(* IEC 61131-3 sources: Palletizer_Control_with_Automation_Studio/Palletizer/Logical/Libraries/MTBasics, 3 files *)

(* ---- MTBasics.typ ---- *)
TYPE
	MTBasicsDT1InternalType : 	STRUCT  (*Internal variables of function block MTBasicsDT1.*)
		CycleTime : REAL; (*Task cycle time. Unit: [µs].*)
		ParametersValid : BOOL; (*Data for internal use.*)
		Gain : REAL; (*Data for internal use.*)
		TimeConstant : REAL; (*Data for internal use.*)
		Numerator : ARRAY[0..1]OF LREAL; (*Data for internal use.*)
		Denominator : ARRAY[0..1]OF LREAL; (*Data for internal use.*)
		BVector : ARRAY[0..1]OF LREAL; (*Data for internal use.*)
		AVector : ARRAY[0..1]OF LREAL; (*Data for internal use.*)
		XVector : ARRAY[0..1]OF LREAL; (*Data for internal use.*)
		PresetOK : BOOL; (*Data for internal use.*)
		PresetCoefficients : LREAL; (*Data for internal use.*)
		InOld : REAL; (*Data for internal use.*)
		UpdateOld : BOOL; (*Data for internal use.*)
		EnableOld : BOOL; (*Data for internal use.*)
		EnableDone : BOOL; (*Data for internal use.*)
		DisabledBusy : BOOL; (*Data for internal use.*)
		CounterOld : UDINT; (*Data for internal use.*)
		SysRefParaNew : BOOL; (*Data for internal use.*)
		SystemReference : MTTransferFcnType; (*Data for internal use.*)
	END_STRUCT;
	MTBasicsDT2InternalType : 	STRUCT  (*Internal variables of function block MTBasicsDT2.*)
		CycleTime : REAL; (*Task cycle time. Unit: [µs].*)
		ParametersValid : BOOL; (*Data for internal use.*)
		Gain : REAL; (*Data for internal use.*)
		TimeConstant1 : REAL; (*Data for internal use.*)
		TimeConstant2 : REAL; (*Data for internal use.*)
		Numerator : ARRAY[0..2]OF LREAL; (*Data for internal use.*)
		Denominator : ARRAY[0..2]OF LREAL; (*Data for internal use.*)
		BVector : ARRAY[0..2]OF LREAL; (*Data for internal use.*)
		AVector : ARRAY[0..2]OF LREAL; (*Data for internal use.*)
		XVector : ARRAY[0..1]OF LREAL; (*Data for internal use.*)
		PresetOK : BOOL; (*Data for internal use.*)
		PresetCoefficients : LREAL; (*Data for internal use.*)
		InOld : REAL; (*Data for internal use.*)
		UpdateOld : BOOL; (*Data for internal use.*)
		EnableOld : BOOL; (*Data for internal use.*)
		EnableDone : BOOL; (*Data for internal use.*)
		DisabledBusy : BOOL; (*Data for internal use.*)
		CounterOld : UDINT; (*Data for internal use.*)
		SysRefParaNew : BOOL; (*Data for internal use.*)
		SystemReference : MTTransferFcnType; (*Data for internal use.*)
	END_STRUCT;
	MTBasicsIntegratorInternalType : 	STRUCT  (*Internal variables of function block MTBasicsIntegrator.*)
		CycleTime : REAL; (*Task cycle time. Unit: [s].*)
		ParametersValid : BOOL; (*Data for internal use.*)
		Gain : REAL; (*Data for internal use.*)
		BVector : ARRAY[0..1]OF LREAL; (*Data for internal use.*)
		AVector : ARRAY[0..1]OF LREAL; (*Data for internal use.*)
		XVector : LREAL; (*Data for internal use.*)
		OutPresetValue : REAL; (*Data for internal use.*)
		SetOutOld : BOOL; (*Data for internal use.*)
		UpdateOld : BOOL; (*Data for internal use.*)
		EnableOld : BOOL; (*Data for internal use.*)
		EnableDone : BOOL; (*Data for internal use.*)
		DisabledBusy : BOOL; (*Data for internal use.*)
		CounterOld : UDINT; (*Data for internal use.*)
		SysRefParaNew : BOOL; (*Data for internal use.*)
		SystemReference : MTTransferFcnType; (*Data for internal use.*)
	END_STRUCT;
	MTBasicsLevelCtrlInternalType : 	STRUCT  (*Internal variables of function block MTBasicsLevelController.*)
		CycleTime : REAL; (*Task cycle time. Unit: [s].*)
		ParametersValid : BOOL; (*Data for internal use.*)
		Parameter : MTBasicsLevelCtrlParType; (*Data for internal use.*)
		State : USINT; (*Data for internal use.*)
		UpdateOld : BOOL; (*Data for internal use.*)
		EnableOld : BOOL; (*Data for internal use.*)
	END_STRUCT;
	MTBasicsLevelCtrlParType : 	STRUCT  (*Level controller parameters.*)
		OutputValue1 : REAL; (*1st Output value.*)
		OutputValue2 : REAL; (*2nd Output value.*)
		OutputValue3 : REAL; (*3rd Output value.*)
		ThresholdLevel1 : REAL; (*Threshold level from OutputValue2 to OutputValue1.*)
		ThresholdLevel2 : REAL; (*Threshold level from OutputValue1 to OutputValue2.*)
		ThresholdLevel3 : REAL; (*Threshold level from OutputValue3 to OutputValue2.*)
		ThresholdLevel4 : REAL; (*Threshold level from OutputValue2 to OutputValue3.*)
	END_STRUCT;
	MTBasicsLimiterInternalType : 	STRUCT  (*Internal variables of function block MTBasicsLimiter.*)
		CycleTime : REAL; (*Task cycle time. Unit: [s].*)
		ParametersValid : BOOL; (*Data for internal use.*)
		MaxOut : REAL; (*Data for internal use.*)
		MinOut : REAL; (*Data for internal use.*)
		MaxPosSlewRate : REAL; (*Data for internal use.*)
		MaxNegSlewRate : REAL; (*Data for internal use.*)
		Out : REAL; (*Data for internal use.*)
		OutOld : REAL; (*Data for internal use.*)
		UpperOutLimit : REAL; (*Data for internal use.*)
		LowerOutLimit : REAL; (*Data for internal use.*)
		SetOutOld : BOOL; (*Data for internal use.*)
		UpdateOld : BOOL; (*Data for internal use.*)
		EnableOld : BOOL; (*Data for internal use.*)
	END_STRUCT;
	MTBasicsOscTuningInternalType : 	STRUCT  (*Internal variables of function block MTBasicsOscillationTuning.*)
		CycleTime : REAL; (*Task cycle time. Unit: [s].*)
		ParametersValid : BOOL; (*Data for internal use.*)
		State : USINT; (*State of tuning.*)
		CriticalGain : REAL; (*Critical gain.*)
		OscillationPeriod : REAL; (*Period of oscillation.*)
		NumberOfOscillations : USINT; (*Number of osscilations.*)
		NumberOfPhases : USINT; (*Number of current tuning phase.*)
		MaxRelayOut : REAL; (*Lower limit for output during tuning.*)
		MinRelayOut : REAL; (*Upper limit for output during tuning.*)
		SetValue : REAL; (*Data for internal use.*)
		AverageOutValue : REAL; (*Data for internal use.*)
		MaxActValueTime : ARRAY[0..3]OF REAL; (*Data for internal use.*)
		MinActValueTime : ARRAY[0..3]OF REAL; (*Data for internal use.*)
		MaxActValue : ARRAY[0..3]OF REAL; (*Data for internal use.*)
		MinActValue : ARRAY[0..3]OF REAL; (*Data for internal use.*)
		TuningTime : REAL; (*Data for internal use.*)
		StartingActValue : REAL; (*Data for internal use.*)
		ControlError : REAL; (*Data for internal use.*)
		ActValueAverageAmplitude : REAL; (*Data for internal use.*)
		AverageActValue : REAL; (*Data for internal use.*)
		AverageMaxActValue : REAL; (*Data for internal use.*)
		AverageMinActValue : REAL; (*Data for internal use.*)
		AmplitudeRatio : REAL; (*Data for internal use.*)
		DeltaOut : REAL; (*Data for internal use.*)
		EffectiveDirection : SINT; (*Data for internal use.*)
		StartOld : BOOL; (*Data for internal use.*)
		MinOscillationAmplitude : REAL; (*Data for internal use.*)
		MinOut : REAL; (*Data for internal use.*)
		MaxOut : REAL; (*Data for internal use.*)
		TemporaryQuality : REAL; (*Data for internal use.*)
		TemporaryDerivativeTime : REAL; (*Data for internal use.*)
		TemporaryIntegrationTime : REAL; (*Data for internal use.*)
		TemporaryGain : REAL; (*Data for internal use.*)
		Update : BOOL; (*Data for internal use.*)
		UpdateOld : BOOL; (*Data for internal use.*)
		EnableOld : BOOL; (*Data for internal use.*)
		AverageOutValueSum : REAL; (*Data for internal use.*)
		AverageTime : LREAL; (*Data for internal use.*)
	END_STRUCT;
	MTBasicsPFMInternalType : 	STRUCT  (*Internal variables of function block MTBasicsPFM.*)
		CycleTime : REAL; (*Task cycle time. Unit: [s].*)
		ParametersValid : BOOL; (*Data for internal use.*)
		In : REAL; (*Data for internal use.*)
		PulseWidth : REAL; (*Data for internal use.*)
		MinPause : REAL; (*Data for internal use.*)
		Area : REAL; (*Data for internal use.*)
		AreaC : REAL; (*Data for internal use.*)
		OffTime : REAL; (*Data for internal use.*)
		OnTime : REAL; (*Data for internal use.*)
		Update : BOOL; (*Data for internal use.*)
		UpdateOld : BOOL; (*Data for internal use.*)
		EnableOld : BOOL; (*Data for internal use.*)
	END_STRUCT;
	MTBasicsPIDInternalType : 	STRUCT  (*Internal variables of function block MTBasicsPID.*)
		CycleTime : REAL; (*Task cycle time. Unit: [s].*)
		ParametersValid : BOOL; (*Data for internal use.*)
		PIDParameters : MTPIDParametersType; (*Data for internal use.*)
		MinOut : REAL; (*Data for internal use.*)
		MaxOut : REAL; (*Data for internal use.*)
		Invert : BOOL; (*Data for internal use.*)
		ControlError : REAL; (*Data for internal use.*)
		ControlErrorOld : REAL; (*Data for internal use.*)
		Out : REAL; (*Data for internal use.*)
		HoldIntegration : MTPIDIntegrationEnum; (*Data for internal use.*)
		IntegrationPartPresetValue : REAL; (*Data for internal use.*)
		SetIntegrationPart : BOOL; (*Data for internal use.*)
		SetIntegrationPartOld : BOOL; (*Data for internal use.*)
		EnableTrackingOld : BOOL; (*Data for internal use.*)
		PID_StatusID : DINT; (*Data for internal use.*)
		UpdateOld : BOOL; (*Data for internal use.*)
		EnableOld : BOOL; (*Data for internal use.*)
		EnableDone : BOOL; (*Data for internal use.*)
		DisabledBusy : BOOL; (*Data for internal use.*)
		CounterOld : UDINT; (*Data for internal use.*)
		SysRefParaNew : BOOL; (*Data for internal use.*)
		SystemReference : MTTransferFcnType; (*Data for internal use.*)
	END_STRUCT;
	MTBasicsPT1InternalType : 	STRUCT  (*Internal variables of function block MTBasicsPT1.*)
		CycleTime : REAL; (*Task cycle time. Unit: [s].*)
		ParametersValid : BOOL; (*Data for internal use.*)
		Gain : REAL; (*Data for internal use.*)
		TimeConstant : REAL; (*Data for internal use.*)
		Numerator : ARRAY[0..1]OF LREAL; (*Data for internal use.*)
		Denominator : ARRAY[0..1]OF LREAL; (*Data for internal use.*)
		BVector : ARRAY[0..1]OF LREAL; (*Data for internal use.*)
		AVector : ARRAY[0..1]OF LREAL; (*Data for internal use.*)
		XVector : ARRAY[0..1]OF LREAL; (*Data for internal use.*)
		OutPresetValue : REAL; (*Data for internal use.*)
		PresetCoefficients : LREAL; (*Data for internal use.*)
		PresetOK : BOOL; (*Data for internal use.*)
		SetOutOld : BOOL; (*Data for internal use.*)
		UpdateOld : BOOL; (*Data for internal use.*)
		EnableOld : BOOL; (*Data for internal use.*)
		EnableDone : BOOL; (*Data for internal use.*)
		DisabledBusy : BOOL; (*Data for internal use.*)
		CounterOld : UDINT; (*Data for internal use.*)
		SysRefParaNew : BOOL; (*Data for internal use.*)
		SystemReference : MTTransferFcnType; (*Data for internal use.*)
	END_STRUCT;
	MTBasicsPT2InternalType : 	STRUCT  (*Internal variables of function block MTBasicsPT2.*)
		CycleTime : REAL; (*Task cycle time. Unit: [µs].*)
		ParametersValid : BOOL; (*Data for internal use.*)
		Gain : REAL; (*Data for internal use.*)
		TimeConstant1 : REAL; (*Data for internal use.*)
		TimeConstant2 : REAL; (*Data for internal use.*)
		Numerator : ARRAY[0..2]OF LREAL; (*Data for internal use.*)
		Denominator : ARRAY[0..2]OF LREAL; (*Data for internal use.*)
		BVector : ARRAY[0..2]OF LREAL; (*Data for internal use.*)
		AVector : ARRAY[0..2]OF LREAL; (*Data for internal use.*)
		XVector : ARRAY[0..1]OF LREAL; (*Data for internal use.*)
		OutPresetValue : REAL; (*Data for internal use.*)
		PresetCoefficients : LREAL; (*Data for internal use.*)
		PresetOK : BOOL; (*Data for internal use.*)
		SetOutOld : BOOL; (*Data for internal use.*)
		UpdateOld : BOOL; (*Data for internal use.*)
		EnableOld : BOOL; (*Data for internal use.*)
		EnableDone : BOOL; (*Data for internal use.*)
		DisabledBusy : BOOL; (*Data for internal use.*)
		CounterOld : UDINT; (*Data for internal use.*)
		SysRefParaNew : BOOL; (*Data for internal use.*)
		SystemReference : MTTransferFcnType; (*Data for internal use.*)
	END_STRUCT;
	MTBasicsPWMInternalType : 	STRUCT  (*Internal variables of function block MTBasicsPWM.*)
		CycleTime : REAL; (*Task cycle time. Unit: [s].*)
		ParametersValid : BOOL; (*Data for internal use.*)
		Mode : MTBasicsPWMModeEnum; (*Data for internal use.*)
		MinPulseWidth : REAL; (*Data for internal use.*)
		Period : REAL; (*Data for internal use.*)
		In : REAL; (*Data for internal use.*)
		OnTime : REAL; (*Data for internal use.*)
		OffTime : REAL; (*Data for internal use.*)
		PeriodCounter : REAL; (*Data for internal use.*)
		OnTimeCounter : REAL; (*Data for internal use.*)
		UpdateOld : BOOL; (*Data for internal use.*)
		EnableOld : BOOL; (*Data for internal use.*)
	END_STRUCT;
	MTBasicsPWMModeEnum :
		( (*Pulse mode.*)
		mtBASICS_PULSE_BEGINNING := 0, (*Pulse at the beginning of a period.*)
		mtBASICS_PULSE_MIDDLE := 1 (*Pulse in the middle of a period.*)
		);
	MTBasicsPWMScheduleBufferPtrType : 	STRUCT  (*Buffer pointers of the PWMSchedule.*)
		In : REAL; (*Data for internal use.*)
		OnTime1 : REAL; (*Data for internal use.*)
		OnTime2 : REAL; (*Data for internal use.*)
		OffTime1 : REAL; (*Data for internal use.*)
		OffTime2 : REAL; (*Data for internal use.*)
		OnTimeCounter : REAL; (*Data for internal use.*)
	END_STRUCT;
	MTBasicsPWMScheduleBufferType : 	STRUCT  (*Buffer parameters of the PWMSchedule.*)
		ActIndex : UINT; (*Data for internal use.*)
		ActBufferElements : UINT; (*Data for internal use.*)
		OldBufferElements : {REDUND_UNREPLICABLE} UINT; (*Data for internal use.*)
		PointerTimes : REFERENCE TO MTBasicsPWMScheduleBufferPtrType; (*Data for internal use.*)
		PointerOut : REFERENCE TO BOOL; (*Data for internal use.*)
	END_STRUCT;
	MTBasicsPWMScheduleInternalType : 	STRUCT  (*Internal variables of function block MTBasicsPWM.*)
		CycleTime : REAL; (*Task cycle time. Unit: [s].*)
		ParametersValid : BOOL; (*Data for internal use.*)
		NumberOfInputs : UINT; (*Data for internal use.*)
		Mode : MTBasicsPWMScheduleModeEnum; (*Data for internal use.*)
		MinPulseWidth : REAL; (*Data for internal use.*)
		MinPause : REAL; (*Data for internal use.*)
		Period : REAL; (*Data for internal use.*)
		FreeDutyCycle : REAL; (*Data for internal use.*)
		PeriodCounter : REAL; (*Data for internal use.*)
		Buffer : MTBasicsPWMScheduleBufferType; (*Data for internal use.*)
		UpdateOld : BOOL; (*Data for internal use.*)
		EnableOld : {REDUND_UNREPLICABLE} BOOL; (*Data for internal use.*)
		InhibitUpdate : BOOL; (*Data for internal use.*)
		Update : BOOL; (*Data for internal use.*)
		StatusIDUpdate : DINT; (*Data for internal use.*)
	END_STRUCT;
	MTBasicsPWMScheduleModeEnum :
		( (*Schedule mode.*)
		mtBASICS_SHIFT_PULSE := 0, (*Shift the puls.*)
		mtBASICS_SPLIT_PULSE := 1 (*Split the puls.*)
		);
	MTBasicsStepTuningBufElemType : 	STRUCT  (*Buffer element of MTBasicsStepTuning.*)
		TimeIndex : UDINT; (*Data for internal use.*)
		In : LREAL; (*Data for internal use.*)
		IntIn : LREAL; (*Data for internal use.*)
		IntTimeIn : LREAL; (*Data for internal use.*)
		IntTime2In : LREAL; (*Data for internal use.*)
		Int2In : LREAL; (*Data for internal use.*)
		Int3In : LREAL; (*Data for internal use.*)
		TSum : LREAL; (*Data for internal use.*)
		dTSum : LREAL; (*Data for internal use.*)
		d2TSum : LREAL; (*Data for internal use.*)
		dyACD : LREAL; (*Data for internal use.*)
		d2yACD : LREAL; (*Data for internal use.*)
		d3yACD : LREAL; (*Data for internal use.*)
		DiffIn : LREAL; (*Data for internal use.*)
		Diff2In : LREAL; (*Data for internal use.*)
	END_STRUCT;
	MTBasicsStepTuningInternalType : 	STRUCT  (*Internal variables of function block MTBasicsStepTuning.*)
		CycleTime : REAL; (*Task cycle time. Unit: [s].*)
		ParametersValid : BOOL; (*Data for internal use.*)
		MinActValue : REAL; (*Data for internal use.*)
		MaxActValue : REAL; (*Data for internal use.*)
		MaxTuningTime : REAL; (*Data for internal use.*)
		StepHeight : REAL; (*Data for internal use.*)
		State : MTBasicsStepTuningStateEnum; (*Data for internal use.*)
		TuningTime : REAL; (*Data for internal use.*)
		Area : REAL; (*Data for internal use.*)
		StartActValue : REAL; (*Data for internal use.*)
		SumTime : REAL; (*Data for internal use.*)
		PlantGain : REAL; (*Data for internal use.*)
		LQError : REAL; (*Data for internal use.*)
		LQOutput : ARRAY[0..1]OF REAL; (*Data for internal use.*)
		LQParameterVector : ARRAY[0..2]OF REAL; (*Data for internal use.*)
		ActValueOld : REAL; (*Data for internal use.*)
		SystemSettlingTime : REAL; (*Data for internal use.*)
		SettlingIndex : UINT; (*Data for internal use.*)
		NumberOfSettlingValues : UINT; (*Data for internal use.*)
		NoiseDeadBand : REAL; (*Data for internal use.*)
		StartOld : BOOL; (*Data for internal use.*)
		UpdateOld : BOOL; (*Data for internal use.*)
		EnableOld : BOOL; (*Data for internal use.*)
		Slope : REAL; (*Data for internal use.*)
	END_STRUCT;
	MTBasicsStepTuningStateEnum :
		( (*Tuning state.*)
		mtBASICS_STATE_READY := 1, (*The function block waits for a rising edge of Start.*)
		mtBASICS_STATE_SETTLING := 2, (*It is checked, if the system is in an idle state.*)
		mtBASICS_STATE_STEP := 3, (*The output Out is set to the value StepHeight.*)
		mtBASICS_STATE_CALCULATE_PID := 4 (*PID parameters are calculated.*)
		);
	MTBasicsTimeDelayFcnParaType : 	STRUCT  (*Internal variables for time delay function parameters.*)
		DelayCounter : UDINT; (*Data for internal use.*)
		ActBufferIndex : UDINT; (*Data for internal use.*)
		ActBufferElements : UDINT; (*Data for internal use.*)
		OldBufferElements : UDINT; (*Data for internal use.*)
		DelayTimeAct : REAL; (*Data for internal use.*)
		BufferPointer : REFERENCE TO REAL; (*Data for internal use.*)
	END_STRUCT;
	MTBasicsTimeDelayInternalType : 	STRUCT  (*Internal variables of function block MTBasicsTimeDelay.*)
		CycleTime : REAL; (*Task cycle time. Unit: [s].*)
		DelayTime : REAL; (*Data for internal use.*)
		ParametersValid : BOOL; (*Data for internal use.*)
		InitialValue : REAL; (*Data for internal use.*)
		EnableOld : BOOL; (*Data for internal use.*)
		TimeDelayFcnPara : {REDUND_UNREPLICABLE} MTBasicsTimeDelayFcnParaType; (*Data for internal use.*)
	END_STRUCT;
END_TYPE

(* ---- MTBasics.fun ---- *)
{REDUND_OK} FUNCTION_BLOCK MTBasicsDT1 (*First-order derivative action element.*)
	VAR_INPUT
		Enable : BOOL; (*Enables/Disables the function block.*)
		Gain : REAL; (*Gain factor.*)
		TimeConstant : REAL; (*Time constant. Unit: [s]. Valid value range: TimeConstant >= 0.*)
		Update : BOOL; (*Updates the parameters listed above on a rising edge.*)
		In : REAL; (*Input value.*)
	END_VAR
	VAR_OUTPUT
		Busy : BOOL; (*Function block is busy.*)
		Active : BOOL; (*Function block is active.*)
		Error : BOOL; (*Indicates an error.*)
		StatusID : DINT; (*Status information.*)
		UpdateDone : BOOL; (*Update is done.*)
		Out : REAL; (*Output value.*)
		SystemReference : {REDUND_UNREPLICABLE} UDINT; (*System reference.*)
	END_VAR
	VAR
		Internal : MTBasicsDT1InternalType; (*Data for internal use.*)
	END_VAR
END_FUNCTION_BLOCK

{REDUND_OK} FUNCTION_BLOCK MTBasicsDT2 (*Second-order derivative action element.*)
	VAR_INPUT
		Enable : BOOL; (*Enables/Disables the function block.*)
		Gain : REAL; (*Gain factor.*)
		TimeConstant1 : REAL; (*Time constant. Unit: [s]. Valid value range: TimeConstant1 >= 0.*)
		TimeConstant2 : REAL; (*Time constant. Unit: [s]. Valid value range: TimeConstant2 >= 0.*)
		Update : BOOL; (*Updates the parameters listed above on a rising edge.*)
		In : REAL; (*Input value.*)
	END_VAR
	VAR_OUTPUT
		Busy : BOOL; (*Function block is busy.*)
		Active : BOOL; (*Function block is active.*)
		Error : BOOL; (*Indicates an error.*)
		StatusID : DINT; (*Status information.*)
		UpdateDone : BOOL; (*Update is done.*)
		Out : REAL; (*Output value.*)
		SystemReference : {REDUND_UNREPLICABLE} UDINT; (*System reference.*)
	END_VAR
	VAR
		Internal : MTBasicsDT2InternalType; (*Data for internal use.*)
	END_VAR
END_FUNCTION_BLOCK

{REDUND_OK} FUNCTION_BLOCK MTBasicsIntegrator (*Integrator.*)
	VAR_INPUT
		Enable : BOOL; (*Enables/Disables the function block.*)
		Gain : REAL; (*Gain factor. Valid value range: Gain >= 0.*)
		Update : BOOL; (*Updates the parameters listed above on a rising edge.*)
		In : REAL; (*Input value.*)
		OutPresetValue : REAL; (*Preset value for Out output.*)
		SetOut : BOOL; (*Sets Out to OutPresetValue on rising edge.*)
		HoldOut : BOOL; (*Freezes the function block.*)
	END_VAR
	VAR_OUTPUT
		Busy : BOOL; (*Function block is busy.*)
		Active : BOOL; (*Function block is active.*)
		Error : BOOL; (*Indicates an error.*)
		StatusID : DINT; (*Status information.*)
		UpdateDone : BOOL; (*Update is done.*)
		Out : REAL; (*Output value.*)
		SystemReference : {REDUND_UNREPLICABLE} UDINT; (*System reference.*)
	END_VAR
	VAR
		Internal : MTBasicsIntegratorInternalType; (*Data for internal use.*)
	END_VAR
END_FUNCTION_BLOCK

{REDUND_OK} FUNCTION_BLOCK MTBasicsLevelController (*Level controller.*)
	VAR_INPUT
		Enable : BOOL; (*Enables/Disables the function block.*)
		Parameter : MTBasicsLevelCtrlParType; (*3-step controller parameters.*)
		Update : BOOL; (*Updates the parameters listed above on a rising edge.*)
		In : REAL; (*Input value.*)
	END_VAR
	VAR_OUTPUT
		Active : BOOL; (*Function block is active.*)
		Error : BOOL; (*Indicates an error.*)
		StatusID : DINT; (*Status information.*)
		UpdateDone : BOOL; (*Update is done.*)
		Out : REAL; (*Output value.*)
	END_VAR
	VAR
		Internal : MTBasicsLevelCtrlInternalType; (*Data for internal use.*)
	END_VAR
END_FUNCTION_BLOCK

{REDUND_OK} FUNCTION_BLOCK MTBasicsLimiter (*Limiter.*)
	VAR_INPUT
		Enable : BOOL; (*Enables/Disables the function block.*)
		MinOut : REAL; (*Lower output variable limit. Valid value range: MinOut < MaxOut.*)
		MaxOut : REAL; (*Upper output variable limit. Valid value range: MaxOut > MinOut.*)
		MaxPosSlewRate : REAL; (*Maximum output variable ramp for ramp-up. Unit: [1/s]. Valid value range: MaxPosSlewRate >= 0.*)
		MaxNegSlewRate : REAL; (*Maximum output variable ramp for the ramp-down. Unit: [1/s]. Valid value range: MaxNegSlewRate >= 0.*)
		Update : BOOL; (*Updates the parameters listed above on a rising edge.*)
		In : REAL; (*Input value.*)
		OutPresetValue : REAL; (*Preset value for Out output.*)
		SetOut : BOOL; (*Sets Out to OutPresetValue on rising edge.*)
	END_VAR
	VAR_OUTPUT
		Active : BOOL; (*Function block is active.*)
		Error : BOOL; (*Indicates an error.*)
		StatusID : DINT; (*Status information.*)
		UpdateDone : BOOL; (*Update is done.*)
		Out : REAL; (*Output value.*)
	END_VAR
	VAR
		Internal : MTBasicsLimiterInternalType; (*Data for internal use.*)
	END_VAR
END_FUNCTION_BLOCK

{REDUND_OK} FUNCTION_BLOCK MTBasicsOscillationTuning (*Oscillation tuning for PID.*)
	VAR_INPUT
		Enable : BOOL; (*Enables/Disables the function block.*)
		SetValue : REAL; (*Reference variable (setpoint).*)
		MinOut : REAL; (*Lower manipulated variable limit. Valid value range: MinOut < MaxOut.*)
		MaxOut : REAL; (*Upper manipulated variable limit. Valid value range: MaxOut > MinOut.*)
		Invert : BOOL; (*Inverts the direction of the controller.*)
		Update : BOOL; (*Updates the parameters listed above on a rising edge.*)
		ActValue : REAL; (*Actual measured value.*)
		Start : BOOL; (*Starts the tuning (on positive edge).*)
	END_VAR
	VAR_OUTPUT
		Active : BOOL; (*Function block is active.*)
		Error : BOOL; (*Indicates an error.*)
		StatusID : DINT; (*Status information.*)
		UpdateDone : BOOL; (*Update is done.*)
		Out : REAL; (*Output value (manipulated variable). Value range: MinOut <= Out <= MaxOut.*)
		TuningActive : BOOL; (*Tuning is active.*)
		TuningDone : BOOL; (*Tuning completed.*)
		Quality : REAL; (*Quality of the oscillation tuning. Unit: [%]. Value range: 0 (low) ... 100 (high).*)
		PIDParameters : MTPIDParametersType; (*PID parameters.*)
	END_VAR
	VAR
		Internal : MTBasicsOscTuningInternalType; (*Data for internal use.*)
	END_VAR
END_FUNCTION_BLOCK

{REDUND_OK} FUNCTION_BLOCK MTBasicsPFM (*Pulse frequency modulator.*)
	VAR_INPUT
		Enable : BOOL; (*Enables/Disables the function block.*)
		PulseWidth : REAL; (*Pulse width at the output. Unit: [s]. Valid value range: PulseWidth >= task cycle time.*)
		MinPause : REAL; (*Minimum pause between the pulses at the output. Unit: [s]. Valid value range: MinPause >= task cycle time.*)
		Update : BOOL; (*Updates the parameters listed above on a rising edge.*)
		DutyCycle : REAL; (*Input value.*)
	END_VAR
	VAR_OUTPUT
		Active : BOOL; (*Function block is active.*)
		Error : BOOL; (*Indicates an error.*)
		StatusID : DINT; (*Status information.*)
		UpdateDone : BOOL; (*Update is done.*)
		Out : BOOL; (*Output value.*)
	END_VAR
	VAR
		Internal : MTBasicsPFMInternalType; (*Data for internal use.*)
	END_VAR
END_FUNCTION_BLOCK

{REDUND_OK} FUNCTION_BLOCK MTBasicsPID (*PID controller.*)
	VAR_INPUT
		Enable : BOOL; (*Enables/Disables the function block.*)
		PIDParameters : MTPIDParametersType; (*PID parameters.*)
		MinOut : REAL;
		MaxOut : REAL;
		Invert : BOOL;
		Update : BOOL; (*Updates the parameters listed above on a rising edge.*)
		SetValue : REAL; (*Set value (reference variable).*)
		ActValue : REAL; (*Actual value (controlled variable).*)
		IntegrationPartPresetValue : REAL; (*Preset value for the integral component IntegrationPart.*)
		SetIntegrationPart : BOOL; (*A positive edge on SetIntegrationPart sets the integral component IntegrationPart of the PID controller to IntegrationPartPresetValue.*)
		HoldOut : BOOL; (*Freezes the function block.*)
		TrackingValue : REAL; (*Preset value for the integral component IntegrationPart.*)
		EnableTracking : BOOL; (*A positive edge on SetIntegrationPart sets the integral component IntegrationPart of the PID controller to IntegrationPartPresetValue.*)
		HoldIntegration : MTPIDIntegrationEnum; (*PID parameters.*)
	END_VAR
	VAR_OUTPUT
		Busy : BOOL; (*Function block is busy.*)
		Active : BOOL; (*Function block is active.*)
		Error : BOOL; (*Indicates an error.*)
		StatusID : DINT; (*Status information.*)
		UpdateDone : BOOL; (*Update is done.*)
		Out : REAL; (*Controller output. Value range: MinOut <= Out <= MaxOut.*)
		ControlError : REAL; (*Control error.*)
		ProportionalPart : REAL; (*Proportional component.*)
		IntegrationPart : REAL; (*Integral component.*)
		DerivativePart : REAL; (*Derivative component.*)
		TrackingActive : BOOL; (*Derivative component.*)
		IntegrationStatus : MTPIDIntegrationEnum; (*Derivative component.*)
		SystemReference : {REDUND_UNREPLICABLE} UDINT; (*System reference.*)
	END_VAR
	VAR
		Internal : MTBasicsPIDInternalType; (*Data for internal use.*)
	END_VAR
END_FUNCTION_BLOCK

{REDUND_OK} FUNCTION_BLOCK MTBasicsPT1 (*First-order delay element.*)
	VAR_INPUT
		Enable : BOOL; (*Enables/Disables the function block.*)
		Gain : REAL; (*Gain factor.*)
		TimeConstant : REAL; (*Time constant. Unit: [s]. Valid value range: TimeConstant >= 0.*)
		Update : BOOL; (*Updates the parameters listed above on a rising edge.*)
		In : REAL; (*Input value.*)
		OutPresetValue : REAL; (*Preset value for Out output.*)
		SetOut : BOOL; (*Sets Out to OutPresetValue on rising edge.*)
	END_VAR
	VAR_OUTPUT
		Busy : BOOL; (*Function block is busy.*)
		Active : BOOL; (*Function block is active.*)
		Error : BOOL; (*Indicates an error.*)
		StatusID : DINT; (*Status information.*)
		UpdateDone : BOOL; (*Update is done.*)
		Out : REAL; (*Output value.*)
		SystemReference : {REDUND_UNREPLICABLE} UDINT; (*System reference.*)
	END_VAR
	VAR
		Internal : MTBasicsPT1InternalType; (*Data for internal use.*)
	END_VAR
END_FUNCTION_BLOCK

{REDUND_OK} FUNCTION_BLOCK MTBasicsPT2 (*Second-order delay element.*)
	VAR_INPUT
		Enable : BOOL; (*Enables/Disables the function block.*)
		Gain : REAL; (*Gain.*)
		TimeConstant1 : REAL; (*Time constant. Unit: [s]. Valid value range: TimeConstant1 >= 0.*)
		TimeConstant2 : REAL; (*Time constant. Unit: [s]. Valid value range: TimeConstant2 >= 0.*)
		Update : BOOL; (*Updates the parameters listed above on a rising edge.*)
		In : REAL; (*Input value.*)
		OutPresetValue : REAL; (*Preset value for Out output.*)
		SetOut : BOOL; (*Sets Out to OutPresetValue on rising edge.*)
	END_VAR
	VAR_OUTPUT
		Busy : BOOL; (*Function block is busy.*)
		Active : BOOL; (*Function block is active.*)
		Error : BOOL; (*Indicates an error.*)
		StatusID : DINT; (*Status information.*)
		UpdateDone : BOOL; (*Update is done.*)
		Out : REAL; (*Output value.*)
		SystemReference : {REDUND_UNREPLICABLE} UDINT; (*System reference.*)
	END_VAR
	VAR
		Internal : MTBasicsPT2InternalType; (*Data for internal use.*)
	END_VAR
END_FUNCTION_BLOCK

{REDUND_OK} FUNCTION_BLOCK MTBasicsPWM (*Pulse width modulator.*)
	VAR_INPUT
		Enable : BOOL; (*Enables/Disables the function block.*)
		Mode : MTBasicsPWMModeEnum; (*Pulse mode.*)
		MinPulseWidth : REAL; (*Minimum duration of the output actuator pulses and pauses. Unit: [s]. Valid value range: MinPulseWidth < Period.*)
		Period : REAL; (*Period for the output actuator pulses. Unit: [s]. Valid value range: Period > task cycle time.*)
		Update : BOOL; (*Updates the parameters listed above on a rising edge.*)
		DutyCycle : REAL; (*Input value. Unit: [%]. Valid value range: 0 <= DutyCycle <= 100.*)
	END_VAR
	VAR_OUTPUT
		Active : BOOL; (*Function block is active.*)
		Error : BOOL; (*Indicates an error.*)
		StatusID : DINT; (*Status information.*)
		UpdateDone : BOOL; (*Update is done.*)
		Out : BOOL; (*Output value.*)
	END_VAR
	VAR
		Internal : MTBasicsPWMInternalType; (*Data for internal use.*)
	END_VAR
END_FUNCTION_BLOCK

{REDUND_CONTEXT} FUNCTION_BLOCK MTBasicsPWMSchedule (*Multiple pulse width modulator.*)
	VAR_INPUT
		Enable : BOOL; (*Enables/Disables the function block.*)
		Period : REAL; (*Period for the output actuator pulses. Unit: [s]. Permitted range: Period > Task cycle time.*)
		MinPulseWidth : REAL; (*Minimum duration of the pulses. Unit: [s]. Permitted range: Task cycle time <= MinPulseWidth < Period.*)
		MinPause : REAL; (*Minimum duration of the pauses. Unit: [s]. Permitted range: Task cycle time <= MinPause < Period.*)
		Mode : MTBasicsPWMScheduleModeEnum; (*Pulse mode.*)
		Update : BOOL; (*Updates the parameters listed above on a rising edge.*)
		NumberOfInputs : UINT; (*Number of input signals. Permitted range: 0 < NumberOfInputs <= 500.*)
		DutyCycle : {REDUND_UNREPLICABLE} UDINT; (*Address of an array of real with the iput values. Unit of values of the assigned array: [%].*)
	END_VAR
	VAR_OUTPUT
		Active : BOOL; (*Function block is active.*)
		Error : BOOL; (*Indicates an error.*)
		StatusID : DINT; (*Status information.*)
		UpdateDone : BOOL; (*Update is done.*)
		Out : {REDUND_UNREPLICABLE} UDINT; (*Address for an array of bool with the output values.*)
	END_VAR
	VAR
		Internal : MTBasicsPWMScheduleInternalType; (*Data for internal use.*)
	END_VAR
END_FUNCTION_BLOCK

{REDUND_OK} FUNCTION_BLOCK MTBasicsStepTuning (*Step tuning for PID.*)
	VAR_INPUT
		Enable : BOOL; (*Enables/Disables the function block.*)
		SystemSettlingTime : REAL; (*System settling time.*)
		MaxTuningTime : REAL; (*Maximum tuning time*)
		MinActValue : REAL; (*Minimum value of the controlled variable.*)
		MaxActValue : REAL; (*Maximum value of the controlled variable.*)
		Update : BOOL; (*Updates the parameters listed above on a rising edge.*)
		ActValue : REAL; (*Actual measured value.*)
		StepHeight : REAL; (*Height of step to be applied.*)
		Start : BOOL; (*Starts the tuning (on positive edge).*)
	END_VAR
	VAR_OUTPUT
		Active : BOOL; (*Function block is active.*)
		Error : BOOL; (*Indicates an error.*)
		StatusID : DINT; (*Status information.*)
		UpdateDone : BOOL; (*Update is done.*)
		Out : REAL; (*Output value (manipulated variable). Value range: MinOut <= Out <= MaxOut.*)
		TuningActive : BOOL; (*Tuning is active.*)
		TuningDone : BOOL; (*Tuning completed.*)
		PIDParameters : MTPIDParametersType; (*PID parameters.*)
		Quality : REAL; (*Quality of the step tuning. Unit: [%]. Value range: 0 (low) ... 100 (high).*)
		TuningState : MTBasicsStepTuningStateEnum; (*Current state of the tuning procedure.*)
	END_VAR
	VAR
		Internal : MTBasicsStepTuningInternalType; (*Data for internal use.*)
	END_VAR
END_FUNCTION_BLOCK

{REDUND_CONTEXT} FUNCTION_BLOCK MTBasicsTimeDelay (*Delay element.*)
	VAR_INPUT
		Enable : BOOL; (*Enables/Disables the function block.*)
		DelayTime : REAL; (*Delay time. Unit: [s]. Valid value range: 0 <= DelayTime <= "10000 · task cycle time".*)
		In : REAL; (*Input value.*)
		InitialValue : REAL; (*Initial value for Out output.*)
	END_VAR
	VAR_OUTPUT
		Active : BOOL; (*Function block is active.*)
		Error : BOOL; (*Indicates an error.*)
		StatusID : DINT; (*Status information.*)
		Out : REAL; (*Output value.*)
	END_VAR
	VAR
		Internal : MTBasicsTimeDelayInternalType; (*Data for internal use.*)
	END_VAR
END_FUNCTION_BLOCK

(* ---- MTBasics.var ---- *)
(*Error*)
VAR CONSTANT
	mtBCD_ERR_TIME_CONSTANT1_INVALID : DINT := -1058012139; (*Chosen first time constant is invalid.*)
	mtBCD_ERR_TIME_CONSTANT2_INVALID : DINT := -1058012138; (*Chosen second time constant is invalid.*)
	mtBCD_ERR_THRESHOLD_NOT_DEFINED : DINT := -1058012137; (*Chosen values for the threshold levels are invalid.*)
	mtBCD_ERR_THRESHOLD_INVALID : DINT := -1058012136; (*One of the values for the threshold levels is invalid.*)
	mtBCD_ERR_OUT_VALUE_NOT_DEFINED : DINT := -1058012135; (*Chosen output values are invalid.*)
	mtBCD_ERR_OUTPUT_LIMIT_INVALID : DINT := -1058012134; (*Chosen limitations for output are invalid.*)
	mtBCD_ERR_MAX_POS_SLEW_RATE_NEG : DINT := -1058012133; (*Chosen slew rate for positive direction is invalid.*)
	mtBCD_ERR_MAX_NEG_SLEW_RATE_NEG : DINT := -1058012132; (*Chosen slew rate for negative direction is invalid.*)
	mtBCD_ERR_PULSE_WIDTH_LOW : DINT := -1058012131; (*Chosen pulse width is too low.*)
	mtBCD_ERR_MIN_PAUSE_LOW : DINT := -1058012130; (*The selected minimum pause duration is too low.*)
	mtBCD_ERR_MIN_PULSE_HIGH : DINT := -1058012124; (*The selected minimum pulse duration is too high.*)
	mtBCD_ERR_MIN_PULSE_LOW : DINT := -1058012123; (*The selected minimum pulse duration is too low.*)
	mtBCD_ERR_PERIOD_LOW : DINT := -1058012122; (*The selected period duration is too low.*)
	mtBCD_ERR_NUMBER_OF_INPUTS : DINT := -1058012121; (*The selected number of inputs is invalid.*)
	mtBCD_ERR_SAMPLING_INVALID : DINT := -1058012118; (*The period of the generated oscillation is invalid. *)
	mtBCD_ERR_SETTLING_TIME_INVALID : DINT := -1058012117; (*Chosen duration, in which the settling of the system is detected, is invalid.*)
	mtBCD_ERR_TUNING_TIME_INVALID : DINT := -1058012116; (*Chosen maximum tuning time is invalid.*)
	mtBCD_ERR_ACT_VALUE_NOT_STABLE : DINT := -1058012115; (*The system is not in a settled operating point.*)
	mtBCD_ERR_RANGE_INVALID : DINT := -1058012114; (*Chosen limitations for the input are invalid.*)
	mtBCD_ERR_TUNING_INVALID : DINT := -1058012113; (*Tuning was not successful.*)
	mtBCD_ERR_MIN_PAUSE_HIGH : DINT := -1058012112; (*The selected minimum pause duration is too high.*)
	mtBCD_ERR_MODE_INVALID : DINT := -1058012111; (*The selected mode is invalid.*)
	mtBCD_ERR_NULL_PTR : DINT := -1058012110; (*Null pointer passed to the input.*)
END_VAR
(*Warning*)
VAR CONSTANT
	mtBCD_WRN_TIME_CONSTANT1_INVALID : DINT := -2131753963; (*Chosen first time constant is invalid.*)
	mtBCD_WRN_TIME_CONSTANT2_INVALID : DINT := -2131753962; (*Chosen second time constant is invalid.*)
	mtBCD_WRN_THRESHOLD_NOT_DEFINED : DINT := -2131753961; (*Chosen values for the threshold levels are invalid.*)
	mtBCD_WRN_THRESHOLD_INVALID : DINT := -2131753960; (*One of the values for the threshold levels is invalid.*)
	mtBCD_WRN_OUT_VALUE_NOT_DEFINED : DINT := -2131753959; (*Chosen output values are invalid.*)
	mtBCD_WRN_OUTPUT_LIMIT_INVALID : DINT := -2131753958; (*Chosen limitations for output are invalid.*)
	mtBCD_WRN_MAX_POS_SLEW_RATE_NEG : DINT := -2131753957; (*Chosen slew rate for positive direction is invalid.*)
	mtBCD_WRN_MAX_NEG_SLEW_RATE_NEG : DINT := -2131753956; (*Chosen slew rate for negative direction is invalid.*)
	mtBCD_WRN_PULSE_WIDTH_LOW : DINT := -2131753955; (*Chosen pulse width is too low.*)
	mtBCD_WRN_MIN_PAUSE_LOW : DINT := -2131753954; (*The selected minimum pause duration is too low.*)
	mtBCD_WRN_GAIN_ZERO : DINT := -2131753953; (*Chosen gain is zero.*)
	mtBCD_WRN_FILTER_TIME_LOW : DINT := -2131753948; (*Chosen filter time is invalid.*)
	mtBCD_WRN_MIN_PULSE_HIGH : DINT := -2131753946; (*The selected minimum pulse duration is too high.*)
	mtBCD_WRN_MIN_PULSE_LOW : DINT := -2131753945; (*The selected minimum pulse duration is too low.*)
	mtBCD_WRN_PERIOD_LOW : DINT := -2131753944; (*The selected period duration is too low.*)
	mtBCD_WRN_SETTLING_TIME_INVALID : DINT := -2131753941; (*Chosen duration, in which the settling of the system is detected, is invalid.*)
	mtBCD_WRN_TUNING_TIME_INVALID : DINT := -2131753940; (*Chosen maximum tuning time is invalid.*)
	mtBCD_WRN_STEP_HEIGHT_INVALID : DINT := -2131753939; (*Chosen step height is zero.*)
	mtBCD_WRN_RANGE_INVALID : DINT := -2131753938; (*Chosen limitations for the input are invalid.*)
	mtBCD_WRN_MIN_PAUSE_HIGH : DINT := -2131753937; (*The selected minimum pause duration is too high.*)
	mtBCD_WRN_MODE_INVALID : DINT := -2131753936; (*The selected mode is invalid.*)
END_VAR
(*Information*)
VAR CONSTANT
	mtBCD_INF_TIME_CONSTANT1_ZERO : DINT := 1089471509; (*Operating as P element or PT1 / DT1 element since TimeConstant1 = 0.*)
	mtBCD_INF_TIME_CONSTANT2_ZERO : DINT := 1089471510; (*Operating as P element or PT1 / DT1 element since TimeConstant2 = 0.*)
	mtBCD_INF_TUNING_ABORTED_BY_USER : DINT := 1089471511; (*Tuning aborted by user.*)
END_VAR
